INTERFACE I_SafetyRelay_1

PROPERTY safetyRelayInFault : BOOL
GET
END_GET
END_PROPERTY

END_INTERFACE

(* stored: Version 1.1.0.1, ProductVersion 3.1.4024.12
   Itf I_SafetyRelay_1: Id {1be3e3f9-77e5-4eb1-9303-001e1f4c8386}
   Property safetyRelayInFault: Id {538d14c8-c431-472e-8ae0-5d48da7f3cef}
   Get Get: Id {e19c7ead-4c21-4dda-813f-e77fe8c61248} *)
